// TIA Portal V20 export
TYPE "WT2_Vb_Befehl_UDT"
   STRUCT
      iHandshake : Int;
      Befehl : Struct
         iID : Int;
         iParam : Int;
      END_STRUCT;
      Param : Struct
         dwID : DWord;
         dwValue : DWord;
         iDiv : Int;
         byEditKonfigSet : Byte;
         byReserve : Byte;
         dwReserve2 : DWord;
      END_STRUCT;
      FernVorgabeDig : Struct
         bFernStartbefehl : Bool;
         bSollwertumschAB : Bool;
         b222_Reserve : Bool;
         b223_Reserve : Bool;
         b224_Reserve : Bool;
         b225_Reserve : Bool;
         b226_Reserve : Bool;
         b227_Reserve : Bool;
         by23_Reserve : Byte;
      END_STRUCT;
      rFernSollwert : Real;
      rFernBegrenz : Real;
      rFernLeistungsbeschränkung : Real;
      byReserve : Array[0..28] of Byte;
   END_STRUCT;
END_TYPE
